// TIA Portal V20 export
FUNCTION_BLOCK "PR_TabTrimSeq_Soft2.0 1_workflow_23a3c5"   // FB52, LAD
{ S7_Optimized_Access := 'TRUE' }
// stored: MemoryReserve 100, SetENOAutomatically false
   VAR_INPUT
      iAbort : Bool;
      iAutoRunning : Bool;
      iFaultReset : Bool;
      iPartNotWorkable : Bool;
      iPartWorkable : Bool;
      iRFReadDone : Bool;
      iRFReadError : Bool;
      iRFWriteDone : Bool;
      iRFWriteError : Bool;
      iReject : Bool;
      iReset_fault : Bool;
      iRetry : Bool;
      iRetryCount : Int;
      iSstMode : Bool;
      iSstPB : Bool;
      iStartFrmFibro : Bool;
      iStartFrmFibroSeq : Bool;
      iTrimOver : Bool;
      iZAxisDownOver : Bool;
      iZAxisUpOver : Bool;
   END_VAR
   VAR_OUTPUT
      qError : Array[0..2] of Bool;
      qMessage : Array[0..2] of Bool;
      qScrapSuction : Bool;
      qTrimOprnOver : Bool;
      qTrimStartCmd : Bool;
      qZAxisUp : Bool;
      qzAxisDown : Bool;
   END_VAR
   VAR
      c20_ChkRecovery_T1 : Bool;
      c20_ChkRecovery_T2 : Bool;
      c20_ChkRecovery_T3 : Bool;
      c21_WtRFIDReadOver_T1 : Bool;
      c21_WtRFIDReadOver_T2 : Bool;
      c22_ChkRetryCountRead_T1 : Bool;
      c22_ChkRetryCountRead_T2 : Bool;
      c23_WtOpDecisionRead_T1 : Bool;
      c23_WtOpDecisionRead_T2 : Bool;
      c24_ChkPartWorkable_T1 : Bool;
      c24_ChkPartWorkable_T2 : Bool;
      c61_WtRFIDWriteOver_T1 : Bool;
      c61_WtRFIDWriteOver_T2 : Bool;
      c62_ChkRetryCountWrite_T1 : Bool;
      c62_ChkRetryCountWrite_T2 : Bool;
      c63_WtOpDecisionWrite_T1 : Bool;
      c63_WtOpDecisionWrite_T2 : Bool;
      StateNo : Int;
      s10_WtStart : Bool;
      s10_WtStart_T1 : Bool;
      s1_WtResetRel : Bool;
      s1_WtResetRel_T1 : Bool;
      s20_ChkRecovery : Bool;
      s20_ChkRecovery_T1 : Bool;
      s20_ChkRecovery_T2 : Bool;
      s20_ChkRecovery_T3 : Bool;
      s21_WtRFIDReadOver : Bool;
      s21_WtRFIDReadOver_T1 : Bool;
      s21_WtRFIDReadOver_T2 : Bool;
      s22_ChkRetryCountRead : Bool;
      s22_ChkRetryCountRead_T1 : Bool;
      s22_ChkRetryCountRead_T2 : Bool;
      s23_WtOpDecisionRead : Bool;
      s23_WtOpDecisionRead_T1 : Bool;
      s23_WtOpDecisionRead_T2 : Bool;
      s24_ChkPartWorkable : Bool;
      s24_ChkPartWorkable_T1 : Bool;
      s24_ChkPartWorkable_T2 : Bool;
      s30_WtOperatorAck : Bool;
      s30_WtOperatorAck_T1 : Bool;
      s40_WtZAxisDown : Bool;
      s40_WtZAxisDown_T1 : Bool;
      s50_WtTrimOver : Bool;
      s50_WtTrimOver_T1 : Bool;
      s60_WtZAxisUp : Bool;
      s60_WtZAxisUp_T1 : Bool;
      s61_WtRFIDWriteOver : Bool;
      s61_WtRFIDWriteOver_T1 : Bool;
      s61_WtRFIDWriteOver_T2 : Bool;
      s62_ChkRetryCountWrite : Bool;
      s62_ChkRetryCountWrite_T1 : Bool;
      s62_ChkRetryCountWrite_T2 : Bool;
      s63_WtOpDecisionWrite : Bool;
      s63_WtOpDecisionWrite_T1 : Bool;
      s63_WtOpDecisionWrite_T2 : Bool;
      s70_WtStartLow : Bool;
      s70_WtStartLow_T1 : Bool;
      sAbNormalCond : Bool;
      sRFReadRetryCount : Int;
      sRFWriteRetryCount : Int;
      sSst : Bool;
      sSstPulse : Bool;
      sSstRise : Bool;
      sStWtResetRel : Bool;
      sStWtResetRel_T1 : Bool;
      sTrimProcessActive : Bool;
   END_VAR
   VAR_TEMP
      tOne : Bool;
   END_VAR
   VAR_TEMP   // added for the SCL form of the ladder/FBD networks
      _w1 : Bool;
   END_VAR
BEGIN

REGION Network 1
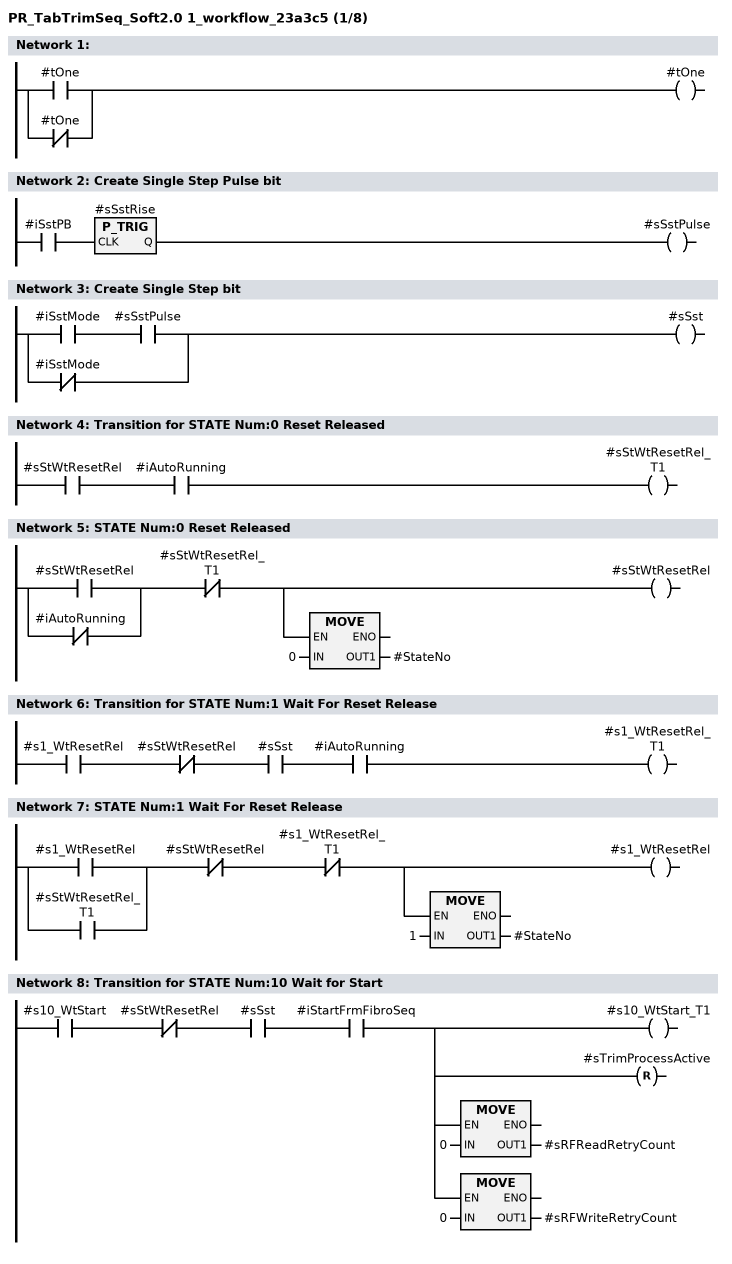
   RUNG wire#powerrail
      Contact( #tOne )
      wire#w1
      Coil( #tOne )
   END_RUNG
   RUNG wire#powerrail
      I_Contact( #tOne )
   END_RUNG wire#w1
   // the same network as SCL:
   #tOne := #tOne OR NOT #tOne;
END_REGION

REGION Network 2: Create Single Step Pulse bit
   RUNG wire#powerrail
      Contact( #iSstPB )
      P_Trig( #sSstRise )
      Coil( #sSstPulse )
   END_RUNG
   // the same network as SCL:
   #_w1 := #iSstPB AND NOT #sSstRise;   // rising edge
   #sSstRise := #iSstPB;
   #sSstPulse := #_w1;
END_REGION

REGION Network 3: Create Single Step bit
   RUNG wire#powerrail
      Contact( #iSstMode )
      Contact( #sSstPulse )
      wire#w1
      Coil( #sSst )
   END_RUNG
   RUNG wire#powerrail
      I_Contact( #iSstMode )
   END_RUNG wire#w1
   // the same network as SCL:
   #sSst := (#iSstMode AND #sSstPulse) OR NOT #iSstMode;
END_REGION

REGION Network 4: Transition for STATE Num:0 Reset Released
   RUNG wire#powerrail
      Contact( #sStWtResetRel )
      Contact( #iAutoRunning )
      Coil( #sStWtResetRel_T1 )
   END_RUNG
   // the same network as SCL:
   #sStWtResetRel_T1 := #sStWtResetRel AND #iAutoRunning;
END_REGION

REGION Network 5: STATE Num:0 Reset Released
   RUNG wire#powerrail
      Contact( #sStWtResetRel )
      wire#w1
      I_Contact( #sStWtResetRel_T1 )
      wire#w2
      Coil( #sStWtResetRel )
   END_RUNG
   RUNG wire#powerrail
      I_Contact( #iAutoRunning )
   END_RUNG wire#w1
   RUNG wire#w2
      { S7_GenerateENO := "TRUE" } Move(in := 0, out1 => #StateNo)
   END_RUNG
   // the same network as SCL:
   #sStWtResetRel := (#sStWtResetRel OR NOT #iAutoRunning) AND NOT #sStWtResetRel_T1;
   IF #sStWtResetRel THEN #StateNo := 0; END_IF;
END_REGION

REGION Network 6: Transition for STATE Num:1 Wait For Reset Release
   RUNG wire#powerrail
      Contact( #s1_WtResetRel )
      I_Contact( #sStWtResetRel )
      Contact( #sSst )
      Contact( #iAutoRunning )
      Coil( #s1_WtResetRel_T1 )
   END_RUNG
   // the same network as SCL:
   #s1_WtResetRel_T1 := #s1_WtResetRel AND NOT #sStWtResetRel AND #sSst AND #iAutoRunning;
END_REGION

REGION Network 7: STATE Num:1 Wait For Reset Release
   RUNG wire#powerrail
      Contact( #s1_WtResetRel )
      wire#w1
      I_Contact( #sStWtResetRel )
      I_Contact( #s1_WtResetRel_T1 )
      wire#w2
      Coil( #s1_WtResetRel )
   END_RUNG
   RUNG wire#powerrail
      Contact( #sStWtResetRel_T1 )
   END_RUNG wire#w1
   RUNG wire#w2
      { S7_GenerateENO := "TRUE" } Move(in := 1, out1 => #StateNo)
   END_RUNG
   // the same network as SCL:
   #s1_WtResetRel := (#s1_WtResetRel OR #sStWtResetRel_T1) AND NOT #sStWtResetRel AND NOT #s1_WtResetRel_T1;
   IF #s1_WtResetRel THEN #StateNo := 1; END_IF;
END_REGION

REGION Network 8: Transition for STATE Num:10 Wait for Start
   RUNG wire#powerrail
      Contact( #s10_WtStart )
      I_Contact( #sStWtResetRel )
      Contact( #sSst )
      Contact( #iStartFrmFibroSeq )
      wire#w1
      Coil( #s10_WtStart_T1 )
   END_RUNG
   RUNG wire#w1
      R_Coil( #sTrimProcessActive )
   END_RUNG
   RUNG wire#w1
      Move(in := 0, out1 => #sRFReadRetryCount)
   END_RUNG
   RUNG wire#w1
      Move(in := 0, out1 => #sRFWriteRetryCount)
   END_RUNG
   // the same network as SCL:
   #s10_WtStart_T1 := #s10_WtStart AND NOT #sStWtResetRel AND #sSst AND #iStartFrmFibroSeq;
   IF #s10_WtStart_T1 THEN
       #sTrimProcessActive := FALSE;
       #sRFReadRetryCount := 0;
       #sRFWriteRetryCount := 0;
   END_IF;
END_REGION

REGION Network 9: STATE Num:10 Wait for Start
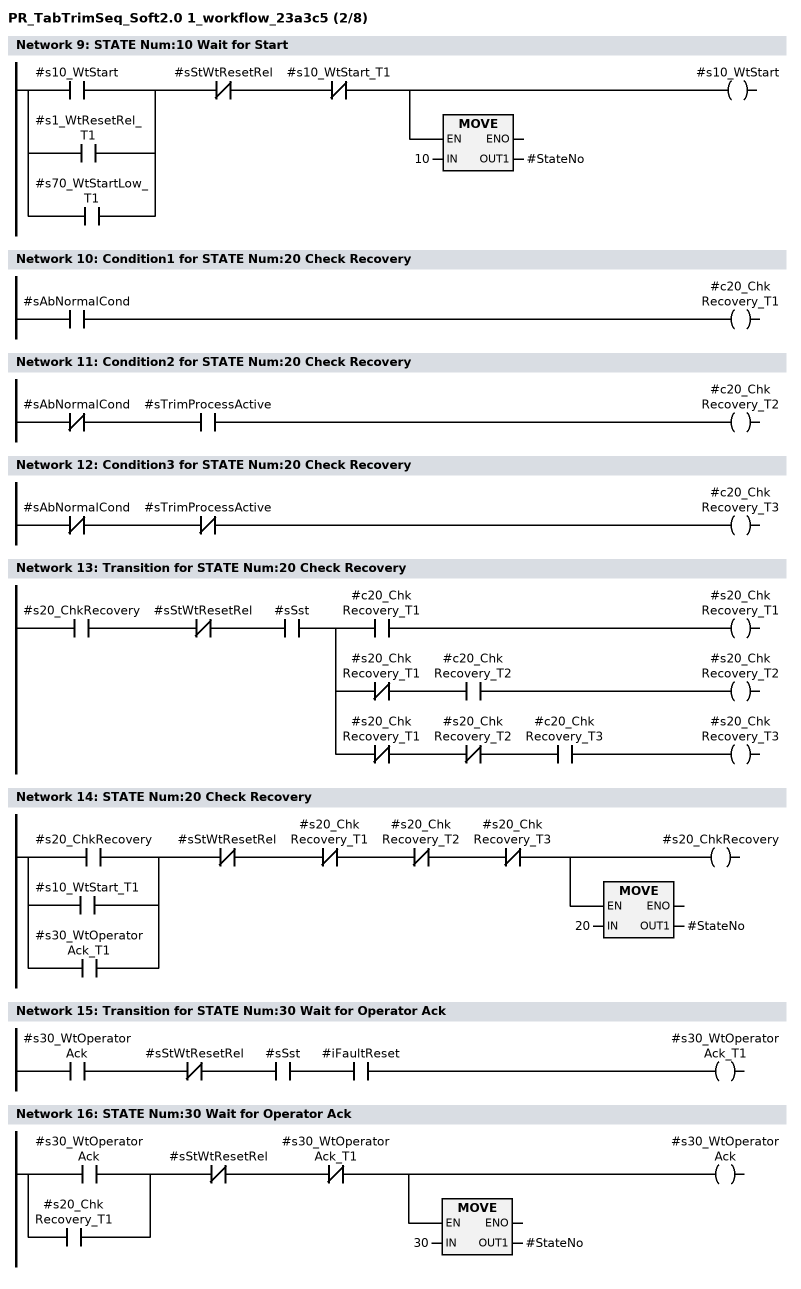
   RUNG wire#powerrail
      Contact( #s10_WtStart )
      wire#w1
      I_Contact( #sStWtResetRel )
      I_Contact( #s10_WtStart_T1 )
      wire#w2
      Coil( #s10_WtStart )
   END_RUNG
   RUNG wire#powerrail
      Contact( #s1_WtResetRel_T1 )
   END_RUNG wire#w1
   RUNG wire#powerrail
      Contact( #s70_WtStartLow_T1 )
   END_RUNG wire#w1
   RUNG wire#w2
      { S7_GenerateENO := "TRUE" } Move(in := 10, out1 => #StateNo)
   END_RUNG
   // the same network as SCL:
   #s10_WtStart := (#s10_WtStart OR #s1_WtResetRel_T1 OR #s70_WtStartLow_T1) AND NOT #sStWtResetRel AND NOT #s10_WtStart_T1;
   IF #s10_WtStart THEN #StateNo := 10; END_IF;
END_REGION

REGION Network 10: Condition1 for STATE Num:20 Check Recovery
   RUNG wire#powerrail
      Contact( #sAbNormalCond )
      Coil( #c20_ChkRecovery_T1 )
   END_RUNG
   // the same network as SCL:
   #c20_ChkRecovery_T1 := #sAbNormalCond;
END_REGION

REGION Network 11: Condition2 for STATE Num:20 Check Recovery
   RUNG wire#powerrail
      I_Contact( #sAbNormalCond )
      Contact( #sTrimProcessActive )
      Coil( #c20_ChkRecovery_T2 )
   END_RUNG
   // the same network as SCL:
   #c20_ChkRecovery_T2 := NOT #sAbNormalCond AND #sTrimProcessActive;
END_REGION

REGION Network 12: Condition3 for STATE Num:20 Check Recovery
   RUNG wire#powerrail
      I_Contact( #sAbNormalCond )
      I_Contact( #sTrimProcessActive )
      Coil( #c20_ChkRecovery_T3 )
   END_RUNG
   // the same network as SCL:
   #c20_ChkRecovery_T3 := NOT #sAbNormalCond AND NOT #sTrimProcessActive;
END_REGION

REGION Network 13: Transition for STATE Num:20 Check Recovery
   RUNG wire#powerrail
      Contact( #s20_ChkRecovery )
      I_Contact( #sStWtResetRel )
      Contact( #sSst )
      wire#w1
      Contact( #c20_ChkRecovery_T1 )
      Coil( #s20_ChkRecovery_T1 )
   END_RUNG
   RUNG wire#w1
      I_Contact( #s20_ChkRecovery_T1 )
      Contact( #c20_ChkRecovery_T2 )
      Coil( #s20_ChkRecovery_T2 )
   END_RUNG
   RUNG wire#w1
      I_Contact( #s20_ChkRecovery_T1 )
      I_Contact( #s20_ChkRecovery_T2 )
      Contact( #c20_ChkRecovery_T3 )
      Coil( #s20_ChkRecovery_T3 )
   END_RUNG
   // the same network as SCL:
   #_w1 := #s20_ChkRecovery AND NOT #sStWtResetRel AND #sSst;
   #s20_ChkRecovery_T1 := #_w1 AND #c20_ChkRecovery_T1;
   #s20_ChkRecovery_T2 := #_w1 AND NOT #s20_ChkRecovery_T1 AND #c20_ChkRecovery_T2;
   #s20_ChkRecovery_T3 := #_w1 AND NOT #s20_ChkRecovery_T1 AND NOT #s20_ChkRecovery_T2 AND #c20_ChkRecovery_T3;
END_REGION

REGION Network 14: STATE Num:20 Check Recovery
   RUNG wire#powerrail
      Contact( #s20_ChkRecovery )
      wire#w1
      I_Contact( #sStWtResetRel )
      I_Contact( #s20_ChkRecovery_T1 )
      I_Contact( #s20_ChkRecovery_T2 )
      I_Contact( #s20_ChkRecovery_T3 )
      wire#w2
      Coil( #s20_ChkRecovery )
   END_RUNG
   RUNG wire#powerrail
      Contact( #s10_WtStart_T1 )
   END_RUNG wire#w1
   RUNG wire#powerrail
      Contact( #s30_WtOperatorAck_T1 )
   END_RUNG wire#w1
   RUNG wire#w2
      { S7_GenerateENO := "TRUE" } Move(in := 20, out1 => #StateNo)
   END_RUNG
   // the same network as SCL:
   #s20_ChkRecovery := (#s20_ChkRecovery OR #s10_WtStart_T1 OR #s30_WtOperatorAck_T1) AND NOT #sStWtResetRel AND NOT #s20_ChkRecovery_T1 AND NOT #s20_ChkRecovery_T2 AND NOT #s20_ChkRecovery_T3;
   IF #s20_ChkRecovery THEN #StateNo := 20; END_IF;
END_REGION

REGION Network 15: Transition for STATE Num:30 Wait for Operator Ack
   RUNG wire#powerrail
      Contact( #s30_WtOperatorAck )
      I_Contact( #sStWtResetRel )
      Contact( #sSst )
      Contact( #iFaultReset )
      Coil( #s30_WtOperatorAck_T1 )
   END_RUNG
   // the same network as SCL:
   #s30_WtOperatorAck_T1 := #s30_WtOperatorAck AND NOT #sStWtResetRel AND #sSst AND #iFaultReset;
END_REGION

REGION Network 16: STATE Num:30 Wait for Operator Ack
   RUNG wire#powerrail
      Contact( #s30_WtOperatorAck )
      wire#w1
      I_Contact( #sStWtResetRel )
      I_Contact( #s30_WtOperatorAck_T1 )
      wire#w2
      Coil( #s30_WtOperatorAck )
   END_RUNG
   RUNG wire#powerrail
      Contact( #s20_ChkRecovery_T1 )
   END_RUNG wire#w1
   RUNG wire#w2
      { S7_GenerateENO := "TRUE" } Move(in := 30, out1 => #StateNo)
   END_RUNG
   // the same network as SCL:
   #s30_WtOperatorAck := (#s30_WtOperatorAck OR #s20_ChkRecovery_T1) AND NOT #sStWtResetRel AND NOT #s30_WtOperatorAck_T1;
   IF #s30_WtOperatorAck THEN #StateNo := 30; END_IF;
END_REGION

REGION Network 17: Actions for STATE Num:30 Wait for Operator Ack
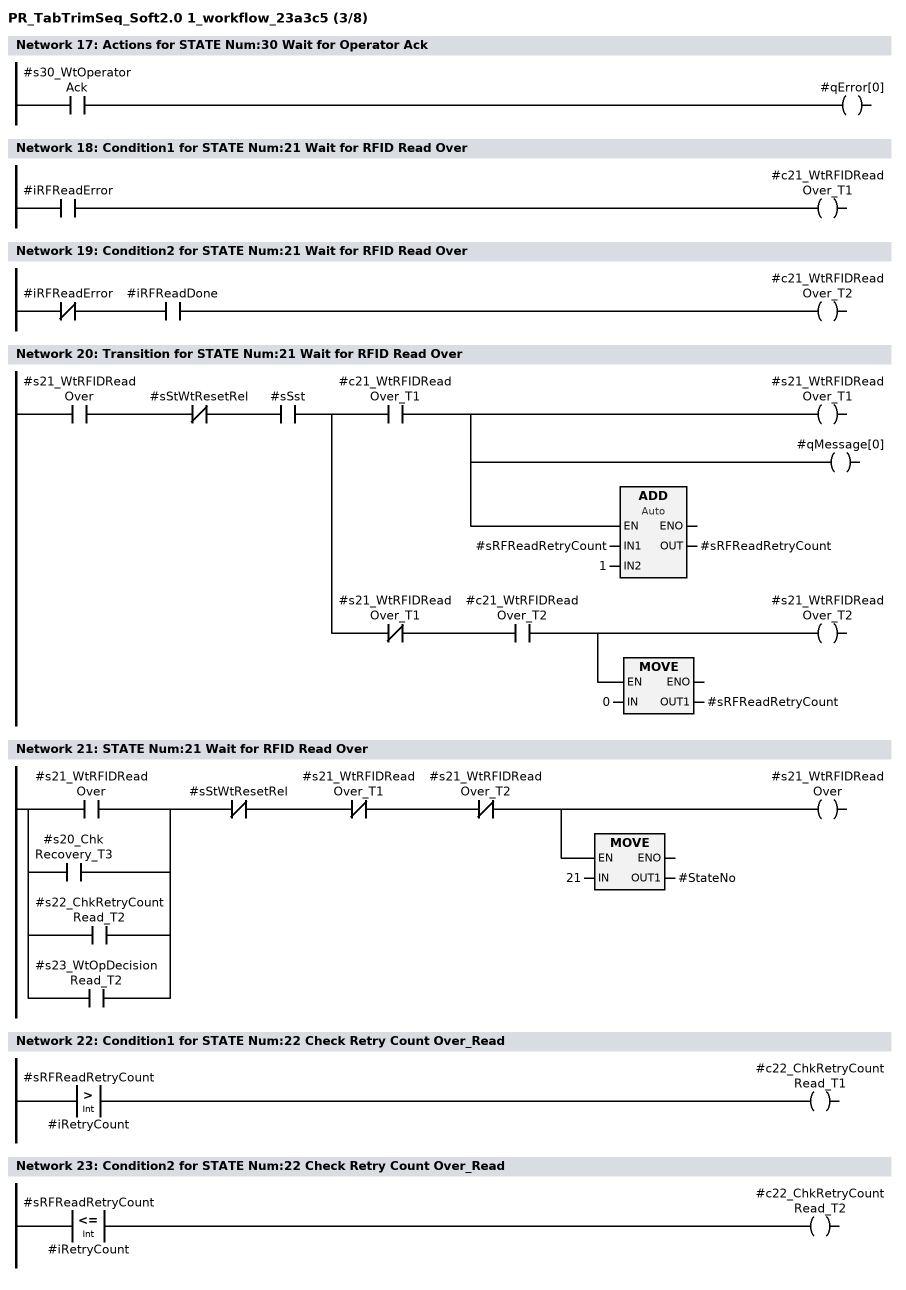
   RUNG wire#powerrail
      Contact( #s30_WtOperatorAck )
      Coil( #qError[0] )
   END_RUNG
   // the same network as SCL:
   #qError[0] := #s30_WtOperatorAck;
END_REGION

REGION Network 18: Condition1 for STATE Num:21 Wait for RFID Read Over
   RUNG wire#powerrail
      Contact( #iRFReadError )
      Coil( #c21_WtRFIDReadOver_T1 )
   END_RUNG
   // the same network as SCL:
   #c21_WtRFIDReadOver_T1 := #iRFReadError;
END_REGION

REGION Network 19: Condition2 for STATE Num:21 Wait for RFID Read Over
   RUNG wire#powerrail
      I_Contact( #iRFReadError )
      Contact( #iRFReadDone )
      Coil( #c21_WtRFIDReadOver_T2 )
   END_RUNG
   // the same network as SCL:
   #c21_WtRFIDReadOver_T2 := NOT #iRFReadError AND #iRFReadDone;
END_REGION

REGION Network 20: Transition for STATE Num:21 Wait for RFID Read Over
   RUNG wire#powerrail
      Contact( #s21_WtRFIDReadOver )
      I_Contact( #sStWtResetRel )
      Contact( #sSst )
      wire#w1
      Contact( #c21_WtRFIDReadOver_T1 )
      wire#w2
      Coil( #s21_WtRFIDReadOver_T1 )
   END_RUNG
   RUNG wire#w2
      Coil( #qMessage[0] )
   END_RUNG
   RUNG wire#w2
      Add(in1 := #sRFReadRetryCount, in2 := 1, out => #sRFReadRetryCount)
   END_RUNG
   RUNG wire#w1
      I_Contact( #s21_WtRFIDReadOver_T1 )
      Contact( #c21_WtRFIDReadOver_T2 )
      wire#w3
      Coil( #s21_WtRFIDReadOver_T2 )
   END_RUNG
   RUNG wire#w3
      Move(in := 0, out1 => #sRFReadRetryCount)
   END_RUNG
   // the same network as SCL:
   #_w1 := #s21_WtRFIDReadOver AND NOT #sStWtResetRel AND #sSst;
   #s21_WtRFIDReadOver_T1 := #_w1 AND #c21_WtRFIDReadOver_T1;
   #qMessage[0] := #s21_WtRFIDReadOver_T1;
   IF #s21_WtRFIDReadOver_T1 THEN #sRFReadRetryCount := #sRFReadRetryCount + 1; END_IF;
   #s21_WtRFIDReadOver_T2 := #_w1 AND NOT #s21_WtRFIDReadOver_T1 AND #c21_WtRFIDReadOver_T2;
   IF #s21_WtRFIDReadOver_T2 THEN #sRFReadRetryCount := 0; END_IF;
END_REGION

REGION Network 21: STATE Num:21 Wait for RFID Read Over
   RUNG wire#powerrail
      Contact( #s21_WtRFIDReadOver )
      wire#w1
      I_Contact( #sStWtResetRel )
      I_Contact( #s21_WtRFIDReadOver_T1 )
      I_Contact( #s21_WtRFIDReadOver_T2 )
      wire#w2
      Coil( #s21_WtRFIDReadOver )
   END_RUNG
   RUNG wire#powerrail
      Contact( #s20_ChkRecovery_T3 )
   END_RUNG wire#w1
   RUNG wire#powerrail
      Contact( #s22_ChkRetryCountRead_T2 )
   END_RUNG wire#w1
   RUNG wire#powerrail
      Contact( #s23_WtOpDecisionRead_T2 )
   END_RUNG wire#w1
   RUNG wire#w2
      { S7_GenerateENO := "TRUE" } Move(in := 21, out1 => #StateNo)
   END_RUNG
   // the same network as SCL:
   #s21_WtRFIDReadOver := (#s21_WtRFIDReadOver OR #s20_ChkRecovery_T3 OR #s22_ChkRetryCountRead_T2 OR #s23_WtOpDecisionRead_T2) AND NOT #sStWtResetRel AND NOT #s21_WtRFIDReadOver_T1 AND NOT #s21_WtRFIDReadOver_T2;
   IF #s21_WtRFIDReadOver THEN #StateNo := 21; END_IF;
END_REGION

REGION Network 22: Condition1 for STATE Num:22 Check Retry Count Over_Read
   RUNG wire#powerrail
      { S7_Templates := "SrcType := Int" } GT_Contact(in1 := #sRFReadRetryCount, in2 := #iRetryCount)
      Coil( #c22_ChkRetryCountRead_T1 )
   END_RUNG
   // the same network as SCL:
   #c22_ChkRetryCountRead_T1 := #sRFReadRetryCount > #iRetryCount;
END_REGION

REGION Network 23: Condition2 for STATE Num:22 Check Retry Count Over_Read
   RUNG wire#powerrail
      { S7_Templates := "SrcType := Int" } LE_Contact(in1 := #sRFReadRetryCount, in2 := #iRetryCount)
      Coil( #c22_ChkRetryCountRead_T2 )
   END_RUNG
   // the same network as SCL:
   #c22_ChkRetryCountRead_T2 := #sRFReadRetryCount <= #iRetryCount;
END_REGION

REGION Network 24: Transition for STATE Num:22 Check Retry Count Over_Read
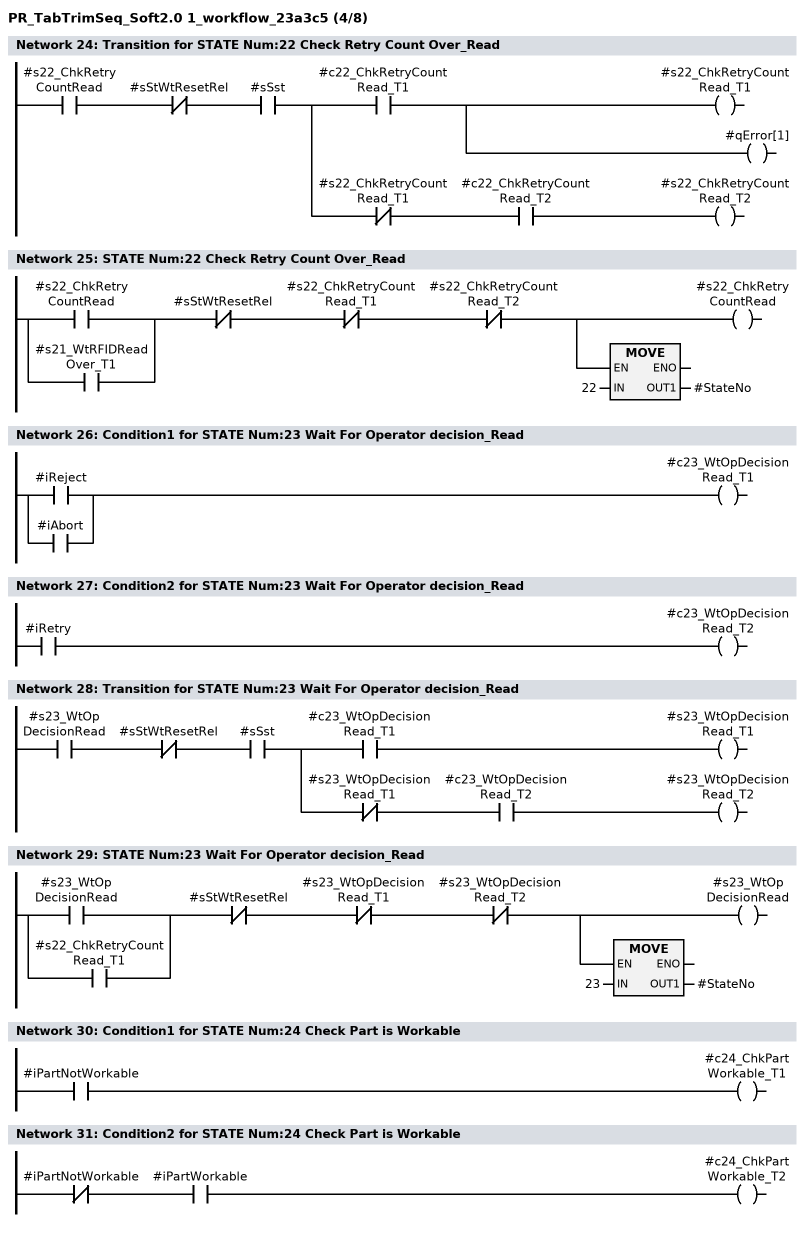
   RUNG wire#powerrail
      Contact( #s22_ChkRetryCountRead )
      I_Contact( #sStWtResetRel )
      Contact( #sSst )
      wire#w1
      Contact( #c22_ChkRetryCountRead_T1 )
      wire#w2
      Coil( #s22_ChkRetryCountRead_T1 )
   END_RUNG
   RUNG wire#w2
      Coil( #qError[1] )
   END_RUNG
   RUNG wire#w1
      I_Contact( #s22_ChkRetryCountRead_T1 )
      Contact( #c22_ChkRetryCountRead_T2 )
      Coil( #s22_ChkRetryCountRead_T2 )
   END_RUNG
   // the same network as SCL:
   #_w1 := #s22_ChkRetryCountRead AND NOT #sStWtResetRel AND #sSst;
   #s22_ChkRetryCountRead_T1 := #_w1 AND #c22_ChkRetryCountRead_T1;
   #qError[1] := #s22_ChkRetryCountRead_T1;
   #s22_ChkRetryCountRead_T2 := #_w1 AND NOT #s22_ChkRetryCountRead_T1 AND #c22_ChkRetryCountRead_T2;
END_REGION

REGION Network 25: STATE Num:22 Check Retry Count Over_Read
   RUNG wire#powerrail
      Contact( #s22_ChkRetryCountRead )
      wire#w1
      I_Contact( #sStWtResetRel )
      I_Contact( #s22_ChkRetryCountRead_T1 )
      I_Contact( #s22_ChkRetryCountRead_T2 )
      wire#w2
      Coil( #s22_ChkRetryCountRead )
   END_RUNG
   RUNG wire#powerrail
      Contact( #s21_WtRFIDReadOver_T1 )
   END_RUNG wire#w1
   RUNG wire#w2
      { S7_GenerateENO := "TRUE" } Move(in := 22, out1 => #StateNo)
   END_RUNG
   // the same network as SCL:
   #s22_ChkRetryCountRead := (#s22_ChkRetryCountRead OR #s21_WtRFIDReadOver_T1) AND NOT #sStWtResetRel AND NOT #s22_ChkRetryCountRead_T1 AND NOT #s22_ChkRetryCountRead_T2;
   IF #s22_ChkRetryCountRead THEN #StateNo := 22; END_IF;
END_REGION

REGION Network 26: Condition1 for STATE Num:23 Wait For Operator decision_Read
   RUNG wire#powerrail
      Contact( #iReject )
      wire#w1
      Coil( #c23_WtOpDecisionRead_T1 )
   END_RUNG
   RUNG wire#powerrail
      Contact( #iAbort )
   END_RUNG wire#w1
   // the same network as SCL:
   #c23_WtOpDecisionRead_T1 := #iReject OR #iAbort;
END_REGION

REGION Network 27: Condition2 for STATE Num:23 Wait For Operator decision_Read
   RUNG wire#powerrail
      Contact( #iRetry )
      Coil( #c23_WtOpDecisionRead_T2 )
   END_RUNG
   // the same network as SCL:
   #c23_WtOpDecisionRead_T2 := #iRetry;
END_REGION

REGION Network 28: Transition for STATE Num:23 Wait For Operator decision_Read
   RUNG wire#powerrail
      Contact( #s23_WtOpDecisionRead )
      I_Contact( #sStWtResetRel )
      Contact( #sSst )
      wire#w1
      Contact( #c23_WtOpDecisionRead_T1 )
      Coil( #s23_WtOpDecisionRead_T1 )
   END_RUNG
   RUNG wire#w1
      I_Contact( #s23_WtOpDecisionRead_T1 )
      Contact( #c23_WtOpDecisionRead_T2 )
      Coil( #s23_WtOpDecisionRead_T2 )
   END_RUNG
   // the same network as SCL:
   #_w1 := #s23_WtOpDecisionRead AND NOT #sStWtResetRel AND #sSst;
   #s23_WtOpDecisionRead_T1 := #_w1 AND #c23_WtOpDecisionRead_T1;
   #s23_WtOpDecisionRead_T2 := #_w1 AND NOT #s23_WtOpDecisionRead_T1 AND #c23_WtOpDecisionRead_T2;
END_REGION

REGION Network 29: STATE Num:23 Wait For Operator decision_Read
   RUNG wire#powerrail
      Contact( #s23_WtOpDecisionRead )
      wire#w1
      I_Contact( #sStWtResetRel )
      I_Contact( #s23_WtOpDecisionRead_T1 )
      I_Contact( #s23_WtOpDecisionRead_T2 )
      wire#w2
      Coil( #s23_WtOpDecisionRead )
   END_RUNG
   RUNG wire#powerrail
      Contact( #s22_ChkRetryCountRead_T1 )
   END_RUNG wire#w1
   RUNG wire#w2
      { S7_GenerateENO := "TRUE" } Move(in := 23, out1 => #StateNo)
   END_RUNG
   // the same network as SCL:
   #s23_WtOpDecisionRead := (#s23_WtOpDecisionRead OR #s22_ChkRetryCountRead_T1) AND NOT #sStWtResetRel AND NOT #s23_WtOpDecisionRead_T1 AND NOT #s23_WtOpDecisionRead_T2;
   IF #s23_WtOpDecisionRead THEN #StateNo := 23; END_IF;
END_REGION

REGION Network 30: Condition1 for STATE Num:24 Check Part is Workable
   RUNG wire#powerrail
      Contact( #iPartNotWorkable )
      Coil( #c24_ChkPartWorkable_T1 )
   END_RUNG
   // the same network as SCL:
   #c24_ChkPartWorkable_T1 := #iPartNotWorkable;
END_REGION

REGION Network 31: Condition2 for STATE Num:24 Check Part is Workable
   RUNG wire#powerrail
      I_Contact( #iPartNotWorkable )
      Contact( #iPartWorkable )
      Coil( #c24_ChkPartWorkable_T2 )
   END_RUNG
   // the same network as SCL:
   #c24_ChkPartWorkable_T2 := NOT #iPartNotWorkable AND #iPartWorkable;
END_REGION

REGION Network 32: Transition for STATE Num:24 Check Part is Workable
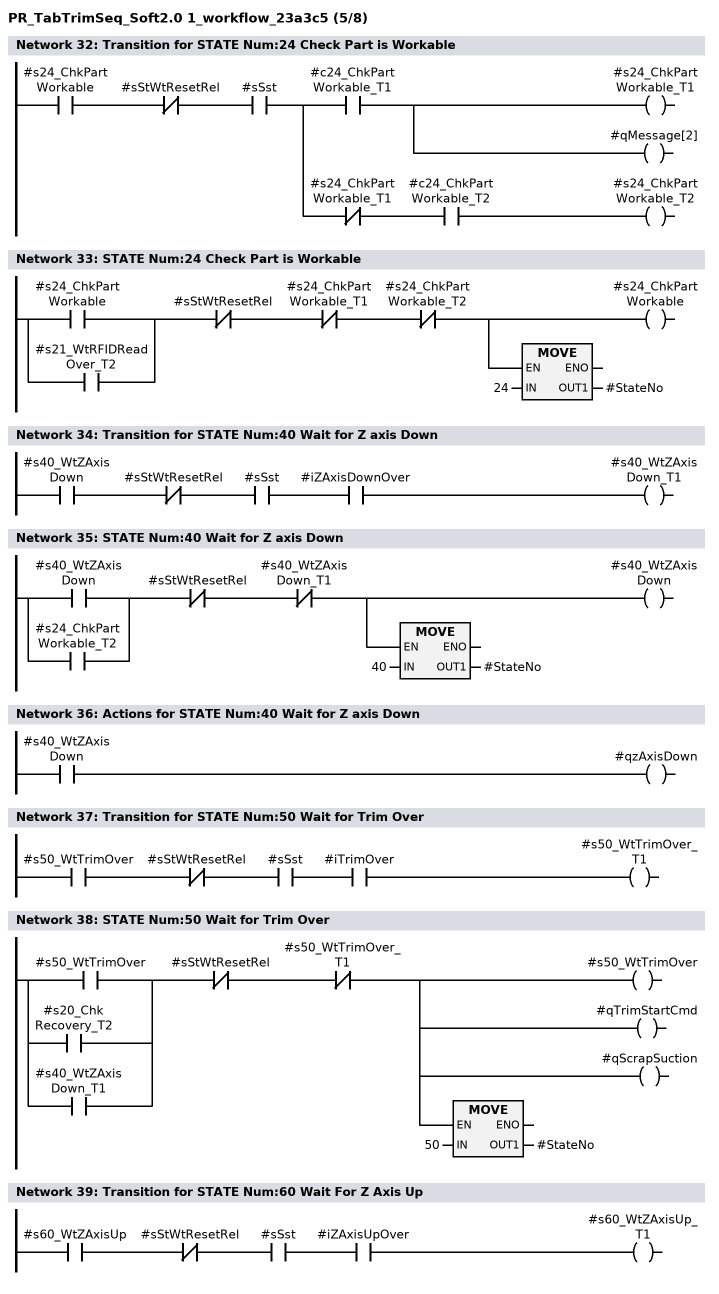
   RUNG wire#powerrail
      Contact( #s24_ChkPartWorkable )
      I_Contact( #sStWtResetRel )
      Contact( #sSst )
      wire#w1
      Contact( #c24_ChkPartWorkable_T1 )
      wire#w2
      Coil( #s24_ChkPartWorkable_T1 )
   END_RUNG
   RUNG wire#w2
      Coil( #qMessage[2] )
   END_RUNG
   RUNG wire#w1
      I_Contact( #s24_ChkPartWorkable_T1 )
      Contact( #c24_ChkPartWorkable_T2 )
      Coil( #s24_ChkPartWorkable_T2 )
   END_RUNG
   // the same network as SCL:
   #_w1 := #s24_ChkPartWorkable AND NOT #sStWtResetRel AND #sSst;
   #s24_ChkPartWorkable_T1 := #_w1 AND #c24_ChkPartWorkable_T1;
   #qMessage[2] := #s24_ChkPartWorkable_T1;
   #s24_ChkPartWorkable_T2 := #_w1 AND NOT #s24_ChkPartWorkable_T1 AND #c24_ChkPartWorkable_T2;
END_REGION

REGION Network 33: STATE Num:24 Check Part is Workable
   RUNG wire#powerrail
      Contact( #s24_ChkPartWorkable )
      wire#w1
      I_Contact( #sStWtResetRel )
      I_Contact( #s24_ChkPartWorkable_T1 )
      I_Contact( #s24_ChkPartWorkable_T2 )
      wire#w2
      Coil( #s24_ChkPartWorkable )
   END_RUNG
   RUNG wire#powerrail
      Contact( #s21_WtRFIDReadOver_T2 )
   END_RUNG wire#w1
   RUNG wire#w2
      { S7_GenerateENO := "TRUE" } Move(in := 24, out1 => #StateNo)
   END_RUNG
   // the same network as SCL:
   #s24_ChkPartWorkable := (#s24_ChkPartWorkable OR #s21_WtRFIDReadOver_T2) AND NOT #sStWtResetRel AND NOT #s24_ChkPartWorkable_T1 AND NOT #s24_ChkPartWorkable_T2;
   IF #s24_ChkPartWorkable THEN #StateNo := 24; END_IF;
END_REGION

REGION Network 34: Transition for STATE Num:40 Wait for Z axis Down
   RUNG wire#powerrail
      Contact( #s40_WtZAxisDown )
      I_Contact( #sStWtResetRel )
      Contact( #sSst )
      Contact( #iZAxisDownOver )
      Coil( #s40_WtZAxisDown_T1 )
   END_RUNG
   // the same network as SCL:
   #s40_WtZAxisDown_T1 := #s40_WtZAxisDown AND NOT #sStWtResetRel AND #sSst AND #iZAxisDownOver;
END_REGION

REGION Network 35: STATE Num:40 Wait for Z axis Down
   RUNG wire#powerrail
      Contact( #s40_WtZAxisDown )
      wire#w1
      I_Contact( #sStWtResetRel )
      I_Contact( #s40_WtZAxisDown_T1 )
      wire#w2
      Coil( #s40_WtZAxisDown )
   END_RUNG
   RUNG wire#powerrail
      Contact( #s24_ChkPartWorkable_T2 )
   END_RUNG wire#w1
   RUNG wire#w2
      { S7_GenerateENO := "TRUE" } Move(in := 40, out1 => #StateNo)
   END_RUNG
   // the same network as SCL:
   #s40_WtZAxisDown := (#s40_WtZAxisDown OR #s24_ChkPartWorkable_T2) AND NOT #sStWtResetRel AND NOT #s40_WtZAxisDown_T1;
   IF #s40_WtZAxisDown THEN #StateNo := 40; END_IF;
END_REGION

REGION Network 36: Actions for STATE Num:40 Wait for Z axis Down
   RUNG wire#powerrail
      Contact( #s40_WtZAxisDown )
      Coil( #qzAxisDown )
   END_RUNG
   // the same network as SCL:
   #qzAxisDown := #s40_WtZAxisDown;
END_REGION

REGION Network 37: Transition for STATE Num:50 Wait for Trim Over
   RUNG wire#powerrail
      Contact( #s50_WtTrimOver )
      I_Contact( #sStWtResetRel )
      Contact( #sSst )
      Contact( #iTrimOver )
      Coil( #s50_WtTrimOver_T1 )
   END_RUNG
   // the same network as SCL:
   #s50_WtTrimOver_T1 := #s50_WtTrimOver AND NOT #sStWtResetRel AND #sSst AND #iTrimOver;
END_REGION

REGION Network 38: STATE Num:50 Wait for Trim Over
   RUNG wire#powerrail
      Contact( #s50_WtTrimOver )
      wire#w1
      I_Contact( #sStWtResetRel )
      I_Contact( #s50_WtTrimOver_T1 )
      wire#w2
      Coil( #s50_WtTrimOver )
   END_RUNG
   RUNG wire#powerrail
      Contact( #s20_ChkRecovery_T2 )
   END_RUNG wire#w1
   RUNG wire#powerrail
      Contact( #s40_WtZAxisDown_T1 )
   END_RUNG wire#w1
   RUNG wire#w2
      Coil( #qTrimStartCmd )
   END_RUNG
   RUNG wire#w2
      Coil( #qScrapSuction )
   END_RUNG
   RUNG wire#w2
      { S7_GenerateENO := "TRUE" } Move(in := 50, out1 => #StateNo)
   END_RUNG
   // the same network as SCL:
   #s50_WtTrimOver := (#s50_WtTrimOver OR #s20_ChkRecovery_T2 OR #s40_WtZAxisDown_T1) AND NOT #sStWtResetRel AND NOT #s50_WtTrimOver_T1;
   #qTrimStartCmd := #s50_WtTrimOver;
   #qScrapSuction := #s50_WtTrimOver;
   IF #s50_WtTrimOver THEN #StateNo := 50; END_IF;
END_REGION

REGION Network 39: Transition for STATE Num:60 Wait For Z Axis Up
   RUNG wire#powerrail
      Contact( #s60_WtZAxisUp )
      I_Contact( #sStWtResetRel )
      Contact( #sSst )
      Contact( #iZAxisUpOver )
      Coil( #s60_WtZAxisUp_T1 )
   END_RUNG
   // the same network as SCL:
   #s60_WtZAxisUp_T1 := #s60_WtZAxisUp AND NOT #sStWtResetRel AND #sSst AND #iZAxisUpOver;
END_REGION

REGION Network 40: STATE Num:60 Wait For Z Axis Up
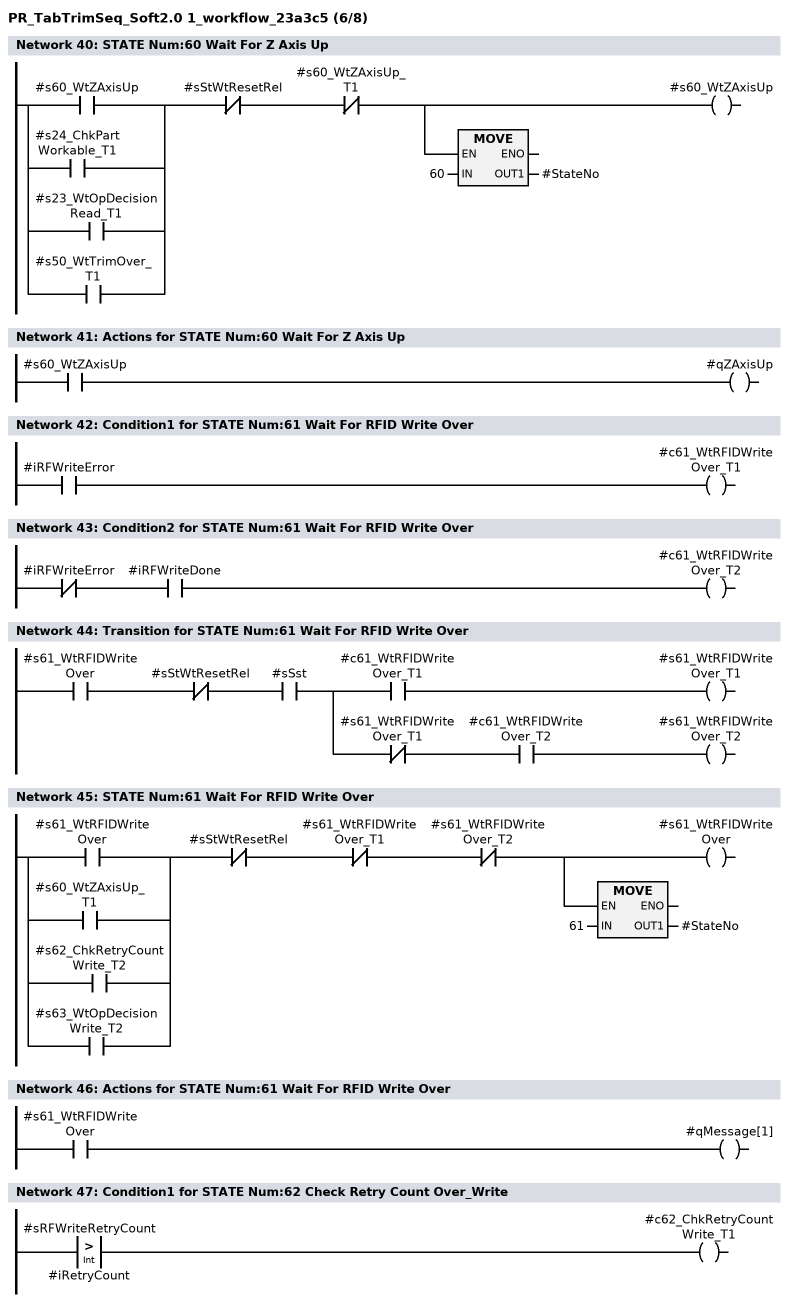
   RUNG wire#powerrail
      Contact( #s60_WtZAxisUp )
      wire#w1
      I_Contact( #sStWtResetRel )
      I_Contact( #s60_WtZAxisUp_T1 )
      wire#w2
      Coil( #s60_WtZAxisUp )
   END_RUNG
   RUNG wire#powerrail
      Contact( #s24_ChkPartWorkable_T1 )
   END_RUNG wire#w1
   RUNG wire#powerrail
      Contact( #s23_WtOpDecisionRead_T1 )
   END_RUNG wire#w1
   RUNG wire#powerrail
      Contact( #s50_WtTrimOver_T1 )
   END_RUNG wire#w1
   RUNG wire#w2
      { S7_GenerateENO := "TRUE" } Move(in := 60, out1 => #StateNo)
   END_RUNG
   // the same network as SCL:
   #s60_WtZAxisUp := (#s60_WtZAxisUp OR #s24_ChkPartWorkable_T1 OR #s23_WtOpDecisionRead_T1 OR #s50_WtTrimOver_T1) AND NOT #sStWtResetRel AND NOT #s60_WtZAxisUp_T1;
   IF #s60_WtZAxisUp THEN #StateNo := 60; END_IF;
END_REGION

REGION Network 41: Actions for STATE Num:60 Wait For Z Axis Up
   RUNG wire#powerrail
      Contact( #s60_WtZAxisUp )
      Coil( #qZAxisUp )
   END_RUNG
   // the same network as SCL:
   #qZAxisUp := #s60_WtZAxisUp;
END_REGION

REGION Network 42: Condition1 for STATE Num:61 Wait For RFID Write Over
   RUNG wire#powerrail
      Contact( #iRFWriteError )
      Coil( #c61_WtRFIDWriteOver_T1 )
   END_RUNG
   // the same network as SCL:
   #c61_WtRFIDWriteOver_T1 := #iRFWriteError;
END_REGION

REGION Network 43: Condition2 for STATE Num:61 Wait For RFID Write Over
   RUNG wire#powerrail
      I_Contact( #iRFWriteError )
      Contact( #iRFWriteDone )
      Coil( #c61_WtRFIDWriteOver_T2 )
   END_RUNG
   // the same network as SCL:
   #c61_WtRFIDWriteOver_T2 := NOT #iRFWriteError AND #iRFWriteDone;
END_REGION

REGION Network 44: Transition for STATE Num:61 Wait For RFID Write Over
   RUNG wire#powerrail
      Contact( #s61_WtRFIDWriteOver )
      I_Contact( #sStWtResetRel )
      Contact( #sSst )
      wire#w1
      Contact( #c61_WtRFIDWriteOver_T1 )
      Coil( #s61_WtRFIDWriteOver_T1 )
   END_RUNG
   RUNG wire#w1
      I_Contact( #s61_WtRFIDWriteOver_T1 )
      Contact( #c61_WtRFIDWriteOver_T2 )
      Coil( #s61_WtRFIDWriteOver_T2 )
   END_RUNG
   // the same network as SCL:
   #_w1 := #s61_WtRFIDWriteOver AND NOT #sStWtResetRel AND #sSst;
   #s61_WtRFIDWriteOver_T1 := #_w1 AND #c61_WtRFIDWriteOver_T1;
   #s61_WtRFIDWriteOver_T2 := #_w1 AND NOT #s61_WtRFIDWriteOver_T1 AND #c61_WtRFIDWriteOver_T2;
END_REGION

REGION Network 45: STATE Num:61 Wait For RFID Write Over
   RUNG wire#powerrail
      Contact( #s61_WtRFIDWriteOver )
      wire#w1
      I_Contact( #sStWtResetRel )
      I_Contact( #s61_WtRFIDWriteOver_T1 )
      I_Contact( #s61_WtRFIDWriteOver_T2 )
      wire#w2
      Coil( #s61_WtRFIDWriteOver )
   END_RUNG
   RUNG wire#powerrail
      Contact( #s60_WtZAxisUp_T1 )
   END_RUNG wire#w1
   RUNG wire#powerrail
      Contact( #s62_ChkRetryCountWrite_T2 )
   END_RUNG wire#w1
   RUNG wire#powerrail
      Contact( #s63_WtOpDecisionWrite_T2 )
   END_RUNG wire#w1
   RUNG wire#w2
      { S7_GenerateENO := "TRUE" } Move(in := 61, out1 => #StateNo)
   END_RUNG
   // the same network as SCL:
   #s61_WtRFIDWriteOver := (#s61_WtRFIDWriteOver OR #s60_WtZAxisUp_T1 OR #s62_ChkRetryCountWrite_T2 OR #s63_WtOpDecisionWrite_T2) AND NOT #sStWtResetRel AND NOT #s61_WtRFIDWriteOver_T1 AND NOT #s61_WtRFIDWriteOver_T2;
   IF #s61_WtRFIDWriteOver THEN #StateNo := 61; END_IF;
END_REGION

REGION Network 46: Actions for STATE Num:61 Wait For RFID Write Over
   RUNG wire#powerrail
      Contact( #s61_WtRFIDWriteOver )
      Coil( #qMessage[1] )
   END_RUNG
   // the same network as SCL:
   #qMessage[1] := #s61_WtRFIDWriteOver;
END_REGION

REGION Network 47: Condition1 for STATE Num:62 Check Retry Count Over_Write
   RUNG wire#powerrail
      { S7_Templates := "SrcType := Int" } GT_Contact(in1 := #sRFWriteRetryCount, in2 := #iRetryCount)
      Coil( #c62_ChkRetryCountWrite_T1 )
   END_RUNG
   // the same network as SCL:
   #c62_ChkRetryCountWrite_T1 := #sRFWriteRetryCount > #iRetryCount;
END_REGION

REGION Network 48: Condition2 for STATE Num:62 Check Retry Count Over_Write
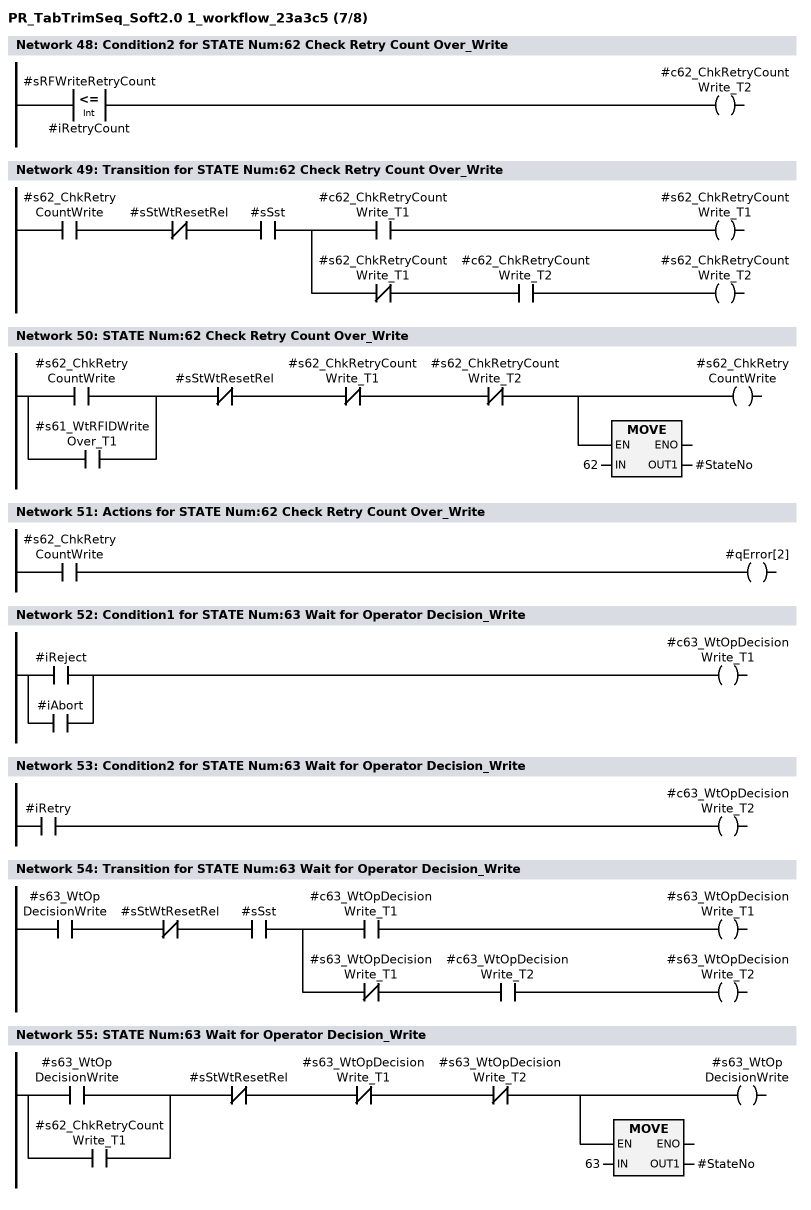
   RUNG wire#powerrail
      { S7_Templates := "SrcType := Int" } LE_Contact(in1 := #sRFWriteRetryCount, in2 := #iRetryCount)
      Coil( #c62_ChkRetryCountWrite_T2 )
   END_RUNG
   // the same network as SCL:
   #c62_ChkRetryCountWrite_T2 := #sRFWriteRetryCount <= #iRetryCount;
END_REGION

REGION Network 49: Transition for STATE Num:62 Check Retry Count Over_Write
   RUNG wire#powerrail
      Contact( #s62_ChkRetryCountWrite )
      I_Contact( #sStWtResetRel )
      Contact( #sSst )
      wire#w1
      Contact( #c62_ChkRetryCountWrite_T1 )
      Coil( #s62_ChkRetryCountWrite_T1 )
   END_RUNG
   RUNG wire#w1
      I_Contact( #s62_ChkRetryCountWrite_T1 )
      Contact( #c62_ChkRetryCountWrite_T2 )
      Coil( #s62_ChkRetryCountWrite_T2 )
   END_RUNG
   // the same network as SCL:
   #_w1 := #s62_ChkRetryCountWrite AND NOT #sStWtResetRel AND #sSst;
   #s62_ChkRetryCountWrite_T1 := #_w1 AND #c62_ChkRetryCountWrite_T1;
   #s62_ChkRetryCountWrite_T2 := #_w1 AND NOT #s62_ChkRetryCountWrite_T1 AND #c62_ChkRetryCountWrite_T2;
END_REGION

REGION Network 50: STATE Num:62 Check Retry Count Over_Write
   RUNG wire#powerrail
      Contact( #s62_ChkRetryCountWrite )
      wire#w1
      I_Contact( #sStWtResetRel )
      I_Contact( #s62_ChkRetryCountWrite_T1 )
      I_Contact( #s62_ChkRetryCountWrite_T2 )
      wire#w2
      Coil( #s62_ChkRetryCountWrite )
   END_RUNG
   RUNG wire#powerrail
      Contact( #s61_WtRFIDWriteOver_T1 )
   END_RUNG wire#w1
   RUNG wire#w2
      { S7_GenerateENO := "TRUE" } Move(in := 62, out1 => #StateNo)
   END_RUNG
   // the same network as SCL:
   #s62_ChkRetryCountWrite := (#s62_ChkRetryCountWrite OR #s61_WtRFIDWriteOver_T1) AND NOT #sStWtResetRel AND NOT #s62_ChkRetryCountWrite_T1 AND NOT #s62_ChkRetryCountWrite_T2;
   IF #s62_ChkRetryCountWrite THEN #StateNo := 62; END_IF;
END_REGION

REGION Network 51: Actions for STATE Num:62 Check Retry Count Over_Write
   RUNG wire#powerrail
      Contact( #s62_ChkRetryCountWrite )
      Coil( #qError[2] )
   END_RUNG
   // the same network as SCL:
   #qError[2] := #s62_ChkRetryCountWrite;
END_REGION

REGION Network 52: Condition1 for STATE Num:63 Wait for Operator Decision_Write
   RUNG wire#powerrail
      Contact( #iReject )
      wire#w1
      Coil( #c63_WtOpDecisionWrite_T1 )
   END_RUNG
   RUNG wire#powerrail
      Contact( #iAbort )
   END_RUNG wire#w1
   // the same network as SCL:
   #c63_WtOpDecisionWrite_T1 := #iReject OR #iAbort;
END_REGION

REGION Network 53: Condition2 for STATE Num:63 Wait for Operator Decision_Write
   RUNG wire#powerrail
      Contact( #iRetry )
      Coil( #c63_WtOpDecisionWrite_T2 )
   END_RUNG
   // the same network as SCL:
   #c63_WtOpDecisionWrite_T2 := #iRetry;
END_REGION

REGION Network 54: Transition for STATE Num:63 Wait for Operator Decision_Write
   RUNG wire#powerrail
      Contact( #s63_WtOpDecisionWrite )
      I_Contact( #sStWtResetRel )
      Contact( #sSst )
      wire#w1
      Contact( #c63_WtOpDecisionWrite_T1 )
      Coil( #s63_WtOpDecisionWrite_T1 )
   END_RUNG
   RUNG wire#w1
      I_Contact( #s63_WtOpDecisionWrite_T1 )
      Contact( #c63_WtOpDecisionWrite_T2 )
      Coil( #s63_WtOpDecisionWrite_T2 )
   END_RUNG
   // the same network as SCL:
   #_w1 := #s63_WtOpDecisionWrite AND NOT #sStWtResetRel AND #sSst;
   #s63_WtOpDecisionWrite_T1 := #_w1 AND #c63_WtOpDecisionWrite_T1;
   #s63_WtOpDecisionWrite_T2 := #_w1 AND NOT #s63_WtOpDecisionWrite_T1 AND #c63_WtOpDecisionWrite_T2;
END_REGION

REGION Network 55: STATE Num:63 Wait for Operator Decision_Write
   RUNG wire#powerrail
      Contact( #s63_WtOpDecisionWrite )
      wire#w1
      I_Contact( #sStWtResetRel )
      I_Contact( #s63_WtOpDecisionWrite_T1 )
      I_Contact( #s63_WtOpDecisionWrite_T2 )
      wire#w2
      Coil( #s63_WtOpDecisionWrite )
   END_RUNG
   RUNG wire#powerrail
      Contact( #s62_ChkRetryCountWrite_T1 )
   END_RUNG wire#w1
   RUNG wire#w2
      { S7_GenerateENO := "TRUE" } Move(in := 63, out1 => #StateNo)
   END_RUNG
   // the same network as SCL:
   #s63_WtOpDecisionWrite := (#s63_WtOpDecisionWrite OR #s62_ChkRetryCountWrite_T1) AND NOT #sStWtResetRel AND NOT #s63_WtOpDecisionWrite_T1 AND NOT #s63_WtOpDecisionWrite_T2;
   IF #s63_WtOpDecisionWrite THEN #StateNo := 63; END_IF;
END_REGION

REGION Network 56: Transition for STATE Num:70 Wait For StartLow
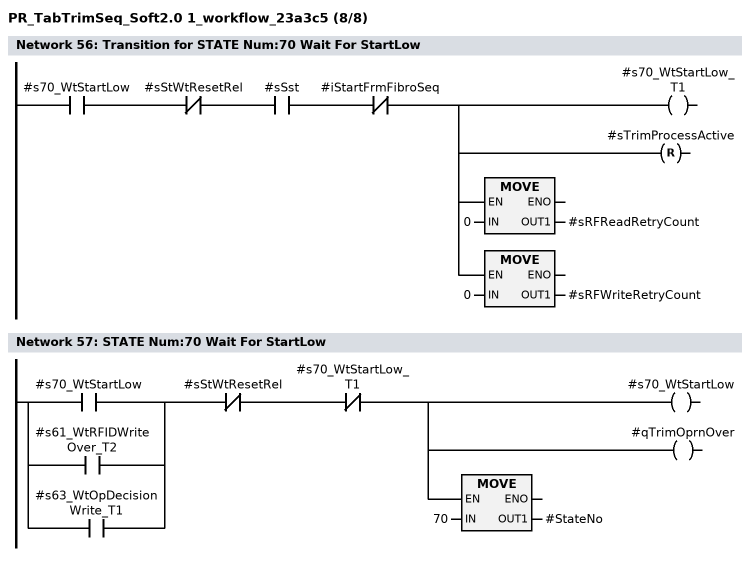
   RUNG wire#powerrail
      Contact( #s70_WtStartLow )
      I_Contact( #sStWtResetRel )
      Contact( #sSst )
      I_Contact( #iStartFrmFibroSeq )
      wire#w1
      Coil( #s70_WtStartLow_T1 )
   END_RUNG
   RUNG wire#w1
      R_Coil( #sTrimProcessActive )
   END_RUNG
   RUNG wire#w1
      Move(in := 0, out1 => #sRFReadRetryCount)
   END_RUNG
   RUNG wire#w1
      Move(in := 0, out1 => #sRFWriteRetryCount)
   END_RUNG
   // the same network as SCL:
   #s70_WtStartLow_T1 := #s70_WtStartLow AND NOT #sStWtResetRel AND #sSst AND NOT #iStartFrmFibroSeq;
   IF #s70_WtStartLow_T1 THEN
       #sTrimProcessActive := FALSE;
       #sRFReadRetryCount := 0;
       #sRFWriteRetryCount := 0;
   END_IF;
END_REGION

REGION Network 57: STATE Num:70 Wait For StartLow
   RUNG wire#powerrail
      Contact( #s70_WtStartLow )
      wire#w1
      I_Contact( #sStWtResetRel )
      I_Contact( #s70_WtStartLow_T1 )
      wire#w2
      Coil( #s70_WtStartLow )
   END_RUNG
   RUNG wire#powerrail
      Contact( #s61_WtRFIDWriteOver_T2 )
   END_RUNG wire#w1
   RUNG wire#powerrail
      Contact( #s63_WtOpDecisionWrite_T1 )
   END_RUNG wire#w1
   RUNG wire#w2
      Coil( #qTrimOprnOver )
   END_RUNG
   RUNG wire#w2
      { S7_GenerateENO := "TRUE" } Move(in := 70, out1 => #StateNo)
   END_RUNG
   // the same network as SCL:
   #s70_WtStartLow := (#s70_WtStartLow OR #s61_WtRFIDWriteOver_T2 OR #s63_WtOpDecisionWrite_T1) AND NOT #sStWtResetRel AND NOT #s70_WtStartLow_T1;
   #qTrimOprnOver := #s70_WtStartLow;
   IF #s70_WtStartLow THEN #StateNo := 70; END_IF;
END_REGION
END_FUNCTION_BLOCK
